// Forçage d'une station (docs/12 § 3)
{attribute 'pack_mode' := '1'}
TYPE ST_StationForce :
STRUCT
    bOutOfProduction : BOOL;
    nReason : USINT;
    tSince : LINT;
    sBy : STRING(24);
END_STRUCT
END_TYPE

(* stored: Version 1.1.0.1, ProductVersion 3.1.4024.12
   DUT ST_StationForce: Id {4a9750ca-8033-505a-bd3f-c011660e65bd} *)
